Fanuc KAREL source: KT00235.KL

PROGRAM KT00235
%NOLOCKGROUP
VAR
  I1: INTEGER
  I2: INTEGER
  OUT: BOOLEAN
BEGIN
  I1 = 2
  I2 = 3
  I1 = 2
  I2 = 3
  OUT = I1 OR I2
END KT00235
